FUNCTION_BLOCK ECController (* EtherCAT master configuration function block *)
  (* Standard: 61499-2; Description: Copyright (c) 2026 Sichuan Qunyuan Technology Co., Ltd. This program and the accompanying materials are made available under the terms of the Eclipse Public License 2.0 which is available at https://www.eclipse.org/legal/epl-2.0/ SPDX-License-Identifier: EPL-2.0 *)
  (* Version 1.1, 2026-10-29, Tim Grocki, Cybernetic Solutions GbR, renamed ControllerIndex to ControllerId to match 4diac FORTE *)
  (* Version 1.0, 2026-04-09, Zijun Tang *)
  PACKAGE eclipse4diac::io::ethercat;
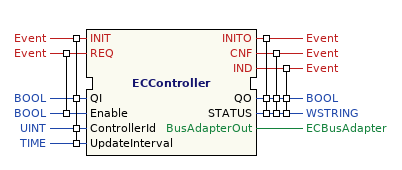
  EVENT_INPUT
    INIT WITH ControllerId, UpdateInterval, QI; (* Initialize the EtherCAT master *)
    REQ WITH Enable; (* Enable or disable cyclic process-data exchange *)
  END_EVENT
  EVENT_OUTPUT
    INITO WITH QO, STATUS; (* Initialization confirm *)
    CNF WITH QO, STATUS; (* Confirmation of the requested enable/disable *)
    IND WITH QO, STATUS; (* Indication of a master or bus state change *)
  END_EVENT
  VAR_INPUT
    QI : BOOL; (* Event input qualifier *)
    Enable : BOOL; (* TRUE starts cyclic EtherCAT I/O *)
    ControllerId : UINT; (* IgH EtherCAT master index *)
    UpdateInterval : TIME := T#1ms; (* Cyclic task period *)
  END_VAR
  VAR_OUTPUT
    QO : BOOL; (* Event output qualifier *)
    STATUS : WSTRING; (* Master status *)
  END_VAR
  PLUGS
    BusAdapterOut : eclipse4diac::io::ethercat::ECBusAdapter; (* Downstream EtherCAT bus adapter *)
  END_PLUGS
END_FUNCTION_BLOCK
